(* PLC project Vn_and2_edit_rename, Beckhoff Automation GmbH TwinCAT PLC Control 3.5.13.21 *)
(* stored: creationDateTime 1970-01-01T00:00:00 *)

PROGRAM Vn_and2_edit_rename

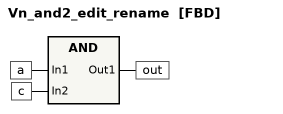
(* FBD diagram, written out as Structured Text *)
out := a AND c;
END_PROGRAM
